SUBAPPLICATION Bool8_TO_logiBUS_QXA8 (* 8 generische digitale Ausgaenge (Kanal frei waehlbar), gemeinsam getriggert durch 1 CNF-Event, adapter-basiert. Generisch fuer jede 8-Bit-Ausgangsgruppe. Schwester-Baustein zu MyLib::sys::Bool8_TO_logiBUS_QX8 (dort logiBUS_QX statt QXA-Adapter). *)
  (* Standard: 61499-2 *)
  (* Version 1.0, 2026-09-09, Franz Höpfinger, Meisterschulen am Ostbahnhof, Angelegt beim Portieren von Uebung_060 nach test_AX zur Wiederverwendung. *)
  PACKAGE MyLib::sys;
  IMPORT logiBUS::io::DQ::logiBUS_DO;
  IMPORT logiBUS::io::DQ::logiBUS_DO_S;
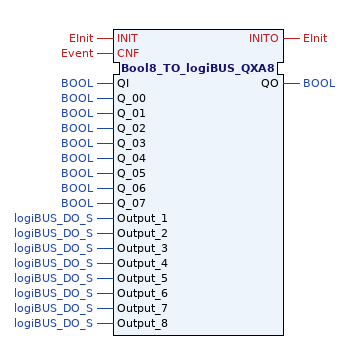
  EVENT_INPUT
    INIT : EInit; (* Initialization Request *)
    CNF;
  END_EVENT
  EVENT_OUTPUT
    INITO : EInit; (* Initialization Confirm *)
  END_EVENT
  VAR_INPUT
    QI : BOOL := TRUE; (* Quality Input - TRUE to enable service *)
    Q_00 : BOOL;
    Q_01 : BOOL;
    Q_02 : BOOL;
    Q_03 : BOOL;
    Q_04 : BOOL;
    Q_05 : BOOL;
    Q_06 : BOOL;
    Q_07 : BOOL;
    Output_1 : logiBUS::io::DQ::logiBUS_DO_S := logiBUS_DO::Invalid; (* Identify the Output Output_Q1..Q8 *)
    Output_2 : logiBUS::io::DQ::logiBUS_DO_S := logiBUS_DO::Invalid; (* Identify the Output Output_Q1..Q8 *)
    Output_3 : logiBUS::io::DQ::logiBUS_DO_S := logiBUS_DO::Invalid; (* Identify the Output Output_Q1..Q8 *)
    Output_4 : logiBUS::io::DQ::logiBUS_DO_S := logiBUS_DO::Invalid; (* Identify the Output Output_Q1..Q8 *)
    Output_5 : logiBUS::io::DQ::logiBUS_DO_S := logiBUS_DO::Invalid; (* Identify the Output Output_Q1..Q8 *)
    Output_6 : logiBUS::io::DQ::logiBUS_DO_S := logiBUS_DO::Invalid; (* Identify the Output Output_Q1..Q8 *)
    Output_7 : logiBUS::io::DQ::logiBUS_DO_S := logiBUS_DO::Invalid; (* Identify the Output Output_Q1..Q8 *)
    Output_8 : logiBUS::io::DQ::logiBUS_DO_S := logiBUS_DO::Invalid; (* Identify the Output Output_Q1..Q8 *)
  END_VAR
  VAR_OUTPUT
    QO : BOOL; (* Quality Output - TRUE if service executed successfully *)
  END_VAR
  FBS
    DigitalOutput_Q4 : logiBUS::io::DQ::logiBUS_QXA;
    DigitalOutput_Q7 : logiBUS::io::DQ::logiBUS_QXA;
    DigitalOutput_Q1 : logiBUS::io::DQ::logiBUS_QXA;
    DigitalOutput_Q5 : logiBUS::io::DQ::logiBUS_QXA;
    DigitalOutput_Q2 : logiBUS::io::DQ::logiBUS_QXA;
    DigitalOutput_Q6 : logiBUS::io::DQ::logiBUS_QXA;
    DigitalOutput_Q8 : logiBUS::io::DQ::logiBUS_QXA;
    DigitalOutput_Q3 : logiBUS::io::DQ::logiBUS_QXA;
    AX_BOOL_TO_X_1 : adapter::conversion::unidirectional::AX_BOOL_TO_X;
    AX_BOOL_TO_X_2 : adapter::conversion::unidirectional::AX_BOOL_TO_X;
    AX_BOOL_TO_X_3 : adapter::conversion::unidirectional::AX_BOOL_TO_X;
    AX_BOOL_TO_X_4 : adapter::conversion::unidirectional::AX_BOOL_TO_X;
    AX_BOOL_TO_X_5 : adapter::conversion::unidirectional::AX_BOOL_TO_X;
    AX_BOOL_TO_X_6 : adapter::conversion::unidirectional::AX_BOOL_TO_X;
    AX_BOOL_TO_X_7 : adapter::conversion::unidirectional::AX_BOOL_TO_X;
    AX_BOOL_TO_X_8 : adapter::conversion::unidirectional::AX_BOOL_TO_X;
    AND_QO : iec61131::booleanOperators::AND_BOOL_8;
  END_FBS
  EVENT_CONNECTIONS
    CNF TO AX_BOOL_TO_X_4.REQ;
    CNF TO AX_BOOL_TO_X_7.REQ;
    CNF TO AX_BOOL_TO_X_1.REQ;
    CNF TO AX_BOOL_TO_X_5.REQ;
    CNF TO AX_BOOL_TO_X_2.REQ;
    CNF TO AX_BOOL_TO_X_6.REQ;
    CNF TO AX_BOOL_TO_X_8.REQ;
    CNF TO AX_BOOL_TO_X_3.REQ;
    INIT TO DigitalOutput_Q4.INIT;
    DigitalOutput_Q4.INITO TO DigitalOutput_Q7.INIT;
    DigitalOutput_Q7.INITO TO DigitalOutput_Q1.INIT;
    DigitalOutput_Q1.INITO TO DigitalOutput_Q5.INIT;
    DigitalOutput_Q5.INITO TO DigitalOutput_Q2.INIT;
    DigitalOutput_Q2.INITO TO DigitalOutput_Q6.INIT;
    DigitalOutput_Q6.INITO TO DigitalOutput_Q8.INIT;
    DigitalOutput_Q8.INITO TO DigitalOutput_Q3.INIT;
    DigitalOutput_Q3.INITO TO INITO;
    DigitalOutput_Q3.INITO TO AND_QO.REQ;
  END_CONNECTIONS
  DATA_CONNECTIONS
    Q_06 TO AX_BOOL_TO_X_7.OUT;
    Q_00 TO AX_BOOL_TO_X_1.OUT;
    Q_04 TO AX_BOOL_TO_X_5.OUT;
    Q_01 TO AX_BOOL_TO_X_2.OUT;
    Q_05 TO AX_BOOL_TO_X_6.OUT;
    Q_02 TO AX_BOOL_TO_X_3.OUT;
    Q_03 TO AX_BOOL_TO_X_4.OUT;
    Q_07 TO AX_BOOL_TO_X_8.OUT;
    Output_1 TO DigitalOutput_Q1.Output;
    Output_2 TO DigitalOutput_Q2.Output;
    Output_3 TO DigitalOutput_Q3.Output;
    Output_4 TO DigitalOutput_Q4.Output;
    Output_5 TO DigitalOutput_Q5.Output;
    Output_6 TO DigitalOutput_Q6.Output;
    Output_7 TO DigitalOutput_Q7.Output;
    Output_8 TO DigitalOutput_Q8.Output;
    QI TO DigitalOutput_Q4.QI;
    QI TO DigitalOutput_Q7.QI;
    QI TO DigitalOutput_Q1.QI;
    QI TO DigitalOutput_Q5.QI;
    QI TO DigitalOutput_Q2.QI;
    QI TO DigitalOutput_Q6.QI;
    QI TO DigitalOutput_Q8.QI;
    QI TO DigitalOutput_Q3.QI;
    DigitalOutput_Q4.QO TO AND_QO.IN1;
    DigitalOutput_Q7.QO TO AND_QO.IN2;
    DigitalOutput_Q1.QO TO AND_QO.IN3;
    DigitalOutput_Q5.QO TO AND_QO.IN4;
    DigitalOutput_Q2.QO TO AND_QO.IN5;
    DigitalOutput_Q6.QO TO AND_QO.IN6;
    DigitalOutput_Q8.QO TO AND_QO.IN7;
    DigitalOutput_Q3.QO TO AND_QO.IN8;
    AND_QO.OUT TO QO;
  END_CONNECTIONS
  ADAPTER_CONNECTIONS
    AX_BOOL_TO_X_1.AX_OUT TO DigitalOutput_Q1.OUT;
    AX_BOOL_TO_X_2.AX_OUT TO DigitalOutput_Q2.OUT;
    AX_BOOL_TO_X_3.AX_OUT TO DigitalOutput_Q3.OUT;
    AX_BOOL_TO_X_4.AX_OUT TO DigitalOutput_Q4.OUT;
    AX_BOOL_TO_X_5.AX_OUT TO DigitalOutput_Q5.OUT;
    AX_BOOL_TO_X_6.AX_OUT TO DigitalOutput_Q6.OUT;
    AX_BOOL_TO_X_7.AX_OUT TO DigitalOutput_Q7.OUT;
    AX_BOOL_TO_X_8.AX_OUT TO DigitalOutput_Q8.OUT;
  END_CONNECTIONS
END_SUBAPPLICATION
